KUKA KRL program: folge11.src, folge11.dat

--- folge11.src ---
&ACCESS RVP
&REL 1
&COMMENT bt2krl vw-ks24 production Folge 11 plan 16#A1BE
DEF FOLGE11()
   ; Generated by bt2krl 0.1.0 from bt2plc plan bt_1792156523_scene_fit (cell scene_fit), PLAN_ID 16#A1BE
   ; Robot robot1 (R1), controller robot1, model unknown, joint mapping identity
   ; Profile vw-ks24 (VW KS24 / TPVW 8.1.8).
   ; Do not edit: regenerate with bt2krl (plain KRL, no inline forms).
   ; Production Folge: 3 ops; per op: P_PktNr_SPS, interlock request + MAKRO20 handshake, motion (exact stop at the end), hold, interlock release
   ; The VW tech package does the Folge handshake (cell.src, AUE_INIT/WAIT/END).
   ;FOLD AUE INIT
      VW(#VW_AUE_INIT,TRUE)
      PENTER:
      INTERRUPT DECL 10 WHEN $CYCFLAG[254]==FALSE DO VW(#FB_STOP,TRUE)
      INTERRUPT ON 10
      INT10=TRUE
   ;ENDFOLD
   ;FOLD VWP0 P0 10 PCT
      ; P0 = home: VW_INIT runs BAS(#INITMOV); AUE_WAIT later sets $H_POS here
      VW(#VW_INIT,TRUE)
      VW_USR_R (#USR_INIT)
      BAS(#VEL_PTP,10)
      $APO.CPTP=100
      PTP P0
      $OUT[15]=TRUE ; PF0 Grundstellung
      ; MAKRO0 RUECKSETZEN_EA: resets A33-A96 (also the tool releases)
      SEL_RES=SELECT(#MAKRO,0,TRUE,,,,,FALSE)
   ;ENDFOLD
   ;FOLD VWAUEWAIT
      VW(#VW_AUE_WAIT,TRUE )
      IF N_VW==TRUE THEN
         GOTO PEXIT
      ENDIF
   ;ENDFOLD
   ;FOLD VWSTART 16#00000003
      ; release every interlock this robot uses: IL01=V1 IL02=V2
      $OUT[15]=FALSE ; PF0 off
      ; MAKRO50 Ini Merker: the cyclic flags of the driving conditions
      SEL_RES=SELECT(#MAKRO,50,TRUE,,,,,FALSE)
      $OUT[41]=TRUE ; release V1
      $OUT[42]=TRUE ; release V2
   ;ENDFOLD
   ;FOLD VWFB 16#00000000
      VALCYCFL30=$CYCFLAG[254]
      $CYCFLAG[254]=($CYCFLAG[30]) AND $CYCFLAG[255] OR ($TIMER[61]<0)
      VW(#FB_CHECK,TRUE)
   ;ENDFOLD
   ;FOLD OP 1 W02 MASK 16#00000001
      ; zones IL01
      P_PktNr_SPS=1
      ;FOLD VWLOCK 16#00000001
         ; enter IL01=V1
         $OUT[81]=TRUE ; request V1
         ; MAKRO20 semantics, inline for these interlocks only
         $OUT[41]=$OUT[41] OR $OUT[81]
         ; PLC grant of the request
         $LOOP_MSG[]="E81"
         $LOOP_CONT=TRUE
         WAIT FOR ($IN[81]) OR (NOT $LOOP_CONT AND ($MODE_OP<>#EX))
         $LOOP_MSG[]="                                                                                                                                "
         ; partner release
         $LOOP_MSG[]="E41"
         $LOOP_CONT=TRUE
         WAIT FOR ($IN[41]) OR (NOT $LOOP_CONT AND ($MODE_OP<>#EX))
         $LOOP_MSG[]="                                                                                                                                "
         $OUT[41]=FALSE ; occupied
         $OUT[81]=FALSE
      ;ENDFOLD
      ;FOLD VWFB 16#00000001
         VALCYCFL30=$CYCFLAG[254]
         $CYCFLAG[254]=($CYCFLAG[30] AND $IN[41]) AND $CYCFLAG[255] OR ($TIMER[61]<0)
         VW(#FB_CHECK,TRUE)
      ;ENDFOLD
      BAS(#VEL_PTP,3)
      PTP P1 C_PTP
      BAS(#VEL_PTP,5)
      PTP P2 C_PTP
      BAS(#VEL_PTP,8)
      PTP P3 C_PTP
      BAS(#VEL_PTP,11)
      PTP P4 C_PTP
      BAS(#VEL_PTP,13)
      PTP P5 C_PTP
      BAS(#VEL_PTP,12)
      PTP P6 C_PTP
      BAS(#VEL_PTP,9)
      PTP P7 C_PTP
      BAS(#VEL_PTP,7)
      PTP P8 C_PTP
      BAS(#VEL_PTP,5)
      PTP P9 C_PTP
      BAS(#VEL_PTP,2)
      PTP P10 C_PTP
      BAS(#VEL_PTP,6)
      PTP P11 C_PTP
      BAS(#VEL_PTP,8)
      PTP P12 C_PTP
      BAS(#VEL_PTP,3)
      PTP P13
      WAIT SEC 0.5 ; hold
      ;FOLD VWUNLOCK 16#00000001
         ; leave IL01=V1
         $OUT[41]=TRUE ; release V1
      ;ENDFOLD
      ;FOLD VWFB 16#00000000
         VALCYCFL30=$CYCFLAG[254]
         $CYCFLAG[254]=($CYCFLAG[30]) AND $CYCFLAG[255] OR ($TIMER[61]<0)
         VW(#FB_CHECK,TRUE)
      ;ENDFOLD
      WAIT SEC 0.1 ; step dwell
   ;ENDFOLD
   ;FOLD OP 2 W04 MASK 16#00000002
      ; zones IL02
      P_PktNr_SPS=2
      ;FOLD VWLOCK 16#00000002
         ; enter IL02=V2
         $OUT[82]=TRUE ; request V2
         ; MAKRO20 semantics, inline for these interlocks only
         $OUT[42]=$OUT[42] OR $OUT[82]
         ; PLC grant of the request
         $LOOP_MSG[]="E82"
         $LOOP_CONT=TRUE
         WAIT FOR ($IN[82]) OR (NOT $LOOP_CONT AND ($MODE_OP<>#EX))
         $LOOP_MSG[]="                                                                                                                                "
         ; partner release
         $LOOP_MSG[]="E42"
         $LOOP_CONT=TRUE
         WAIT FOR ($IN[42]) OR (NOT $LOOP_CONT AND ($MODE_OP<>#EX))
         $LOOP_MSG[]="                                                                                                                                "
         $OUT[42]=FALSE ; occupied
         $OUT[82]=FALSE
      ;ENDFOLD
      ;FOLD VWFB 16#00000002
         VALCYCFL30=$CYCFLAG[254]
         $CYCFLAG[254]=($CYCFLAG[30] AND $IN[42]) AND $CYCFLAG[255] OR ($TIMER[61]<0)
         VW(#FB_CHECK,TRUE)
      ;ENDFOLD
      BAS(#VEL_PTP,4)
      PTP P14 C_PTP
      PTP P15 C_PTP
      BAS(#VEL_PTP,10)
      PTP P16 C_PTP
      BAS(#VEL_PTP,13)
      PTP P17 C_PTP
      BAS(#VEL_PTP,11)
      PTP P18 C_PTP
      BAS(#VEL_PTP,7)
      PTP P19 C_PTP
      BAS(#VEL_PTP,3)
      PTP P20 C_PTP
      BAS(#VEL_PTP,6)
      PTP P21 C_PTP
      BAS(#VEL_PTP,8)
      PTP P22 C_PTP
      BAS(#VEL_PTP,3)
      PTP P23
      WAIT SEC 0.5 ; hold
      ;FOLD VWUNLOCK 16#00000002
         ; leave IL02=V2
         $OUT[42]=TRUE ; release V2
      ;ENDFOLD
      ;FOLD VWFB 16#00000000
         VALCYCFL30=$CYCFLAG[254]
         $CYCFLAG[254]=($CYCFLAG[30]) AND $CYCFLAG[255] OR ($TIMER[61]<0)
         VW(#FB_CHECK,TRUE)
      ;ENDFOLD
      WAIT SEC 0.1 ; step dwell
   ;ENDFOLD
   ;FOLD OP 3 HOME MASK 16#00000001
      ; zones IL01
      P_PktNr_SPS=3
      ;FOLD VWLOCK 16#00000001
         ; enter IL01=V1
         $OUT[81]=TRUE ; request V1
         ; MAKRO20 semantics, inline for these interlocks only
         $OUT[41]=$OUT[41] OR $OUT[81]
         ; PLC grant of the request
         $LOOP_MSG[]="E81"
         $LOOP_CONT=TRUE
         WAIT FOR ($IN[81]) OR (NOT $LOOP_CONT AND ($MODE_OP<>#EX))
         $LOOP_MSG[]="                                                                                                                                "
         ; partner release
         $LOOP_MSG[]="E41"
         $LOOP_CONT=TRUE
         WAIT FOR ($IN[41]) OR (NOT $LOOP_CONT AND ($MODE_OP<>#EX))
         $LOOP_MSG[]="                                                                                                                                "
         $OUT[41]=FALSE ; occupied
         $OUT[81]=FALSE
      ;ENDFOLD
      ;FOLD VWFB 16#00000001
         VALCYCFL30=$CYCFLAG[254]
         $CYCFLAG[254]=($CYCFLAG[30] AND $IN[41]) AND $CYCFLAG[255] OR ($TIMER[61]<0)
         VW(#FB_CHECK,TRUE)
      ;ENDFOLD
      BAS(#VEL_PTP,5)
      PTP P24 C_PTP
      BAS(#VEL_PTP,2)
      PTP P25 C_PTP
      BAS(#VEL_PTP,6)
      PTP P26 C_PTP
      BAS(#VEL_PTP,9)
      PTP P27 C_PTP
      BAS(#VEL_PTP,12)
      PTP P28 C_PTP
      BAS(#VEL_PTP,15)
      PTP P29 C_PTP
      BAS(#VEL_PTP,18)
      PTP P30 C_PTP
      BAS(#VEL_PTP,17)
      PTP P31 C_PTP
      BAS(#VEL_PTP,14)
      PTP P32 C_PTP
      BAS(#VEL_PTP,11)
      PTP P33 C_PTP
      BAS(#VEL_PTP,6)
      PTP P34 C_PTP
      BAS(#VEL_PTP,2)
      PTP P35
      ;FOLD VWMAKRO 15
         ; Gesamtfertigmeldung
         SEL_RES=SELECT(#MAKRO,15,TRUE,,,,,FALSE)
      ;ENDFOLD
      ;FOLD VWUNLOCK 16#00000001
         ; leave IL01=V1
         $OUT[41]=TRUE ; release V1
      ;ENDFOLD
      ;FOLD VWFB 16#00000000
         VALCYCFL30=$CYCFLAG[254]
         $CYCFLAG[254]=($CYCFLAG[30]) AND $CYCFLAG[255] OR ($TIMER[61]<0)
         VW(#FB_CHECK,TRUE)
      ;ENDFOLD
      WAIT SEC 0.1 ; step dwell
   ;ENDFOLD
   P_PktNr_SPS=0
   ;FOLD AUE END
      VW(#VW_AUE_END,TRUE)
      GOTO PENTER
      PEXIT:
   ;ENDFOLD
END

--- folge11.dat ---
&ACCESS RVP
&REL 1
&COMMENT bt2krl vw-ks24 data Folge 11 plan 16#A1BE
DEFDAT FOLGE11
   ; Generated by bt2krl 0.1.0 from bt2plc plan bt_1792156523_scene_fit (cell scene_fit), PLAN_ID 16#A1BE
   ; Robot robot1 (R1), controller robot1, model unknown, joint mapping identity
   ; Profile vw-ks24 (VW KS24 / TPVW 8.1.8).
   ; Do not edit: regenerate with bt2krl (plain KRL, no inline forms).
   EXT BAS (BAS_COMMAND :IN,REAL :IN )
   ; interface to the VW standard routines (as every VW Folge .dat declares them)
   EXT VW (VW_COMMAND :IN,BOOL :IN,REAL :IN,REAL :IN,REAL :IN,REAL :IN,BOOL :IN,E6POS :IN )
   EXT VW_USR_R (VW_USER_CMD :IN,INT :IN,REAL :IN,REAL :IN,REAL :IN,REAL :IN,REAL :IN,REAL :IN,BOOL :IN )
   EXTFCT INT SELECT (SUBTYPE :IN,INT :IN,BOOL :IN,ARI_TYP :IN,INT :IN,BOOL_TYP :IN,INT :IN,BOOL :IN)
   DECL AXIS P0={A1 45.0,A2 -90.0,A3 90.0,A4 0.0,A5 0.0,A6 0.0}
   DECL AXIS P1={A1 43.6012,A2 -89.7676,A3 90.0033,A4 0.0,A5 1.8605,A6 -0.3507}
   DECL AXIS P2={A1 41.9543,A2 -89.4939,A3 90.0071,A4 0.0,A5 4.051,A6 -0.7636}
   DECL AXIS P3={A1 37.1038,A2 -88.6879,A3 90.0185,A4 0.0,A5 10.5026,A6 -1.9796}
   DECL AXIS P4={A1 26.9514,A2 -87.001,A3 90.0423,A4 0.0,A5 24.006,A6 -4.5249}
   DECL AXIS P5={A1 6.8724,A2 -83.6646,A3 90.0893,A4 0.0,A5 50.7127,A6 -9.5588}
   DECL AXIS P6={A1 -4.0921,A2 -81.8426,A3 90.115,A4 0.0,A5 65.2964,A6 -12.3077}
   DECL AXIS P7={A1 -9.8225,A2 -80.8905,A3 90.1284,A4 0.0,A5 72.9183,A6 -13.7444}
   DECL AXIS P8={A1 -12.0109,A2 -80.5268,A3 90.1336,A4 0.0,A5 75.829,A6 -14.293}
   DECL AXIS P9={A1 -14.6956,A2 -80.0807,A3 90.1398,A4 0.0,A5 79.3999,A6 -14.9661}
   DECL AXIS P10={A1 -15.0566,A2 -80.0207,A3 90.1407,A4 0.0,A5 79.88,A6 -15.0566}
   DECL AXIS P11={A1 -15.0566,A2 -79.875,A3 90.7142,A4 0.0,A5 79.1607,A6 -15.0566}
   DECL AXIS P12={A1 -15.0566,A2 -79.6592,A3 91.5498,A4 0.0,A5 78.1094,A6 -15.0566}
   DECL AXIS P13={A1 -15.0566,A2 -78.7933,A3 94.228,A4 0.0,A5 74.5653,A6 -15.0566}
   DECL AXIS P14={A1 -15.0374,A2 -79.913,A3 90.5893,A4 0.0,A5 79.3237,A6 -15.0374}
   DECL AXIS P15={A1 -13.7654,A2 -80.0274,A3 90.142,A4 0.0,A5 79.8854,A6 -13.7654}
   DECL AXIS P16={A1 -9.2939,A2 -80.052,A3 90.1253,A4 0.0,A5 79.9267,A6 -9.2939}
   DECL AXIS P17={A1 8.1168,A2 -80.1118,A3 90.221,A4 0.0,A5 79.8908,A6 8.1168}
   DECL AXIS P18={A1 11.5499,A2 -80.1218,A3 90.2471,A4 0.0,A5 79.8747,A6 11.5498}
   DECL AXIS P19={A1 13.8795,A2 -80.1284,A3 90.2658,A4 0.0,A5 79.8625,A6 13.8794}
   DECL AXIS P20={A1 14.7377,A2 -80.1307,A3 90.273,A4 0.0,A5 79.8577,A6 14.7377}
   DECL AXIS P21={A1 14.7377,A2 -79.9847,A3 90.8466,A4 0.0,A5 79.1381,A6 14.7377}
   DECL AXIS P22={A1 14.7377,A2 -79.7685,A3 91.6823,A4 0.0,A5 78.0862,A6 14.7377}
   DECL AXIS P23={A1 14.7377,A2 -78.9012,A3 94.361,A4 0.0,A5 74.5402,A6 14.7377}
   DECL AXIS P24={A1 14.7377,A2 -79.9556,A3 90.9835,A4 0.0,A5 78.9721,A6 14.7377}
   DECL AXIS P25={A1 15.0076,A2 -80.0451,A3 90.9747,A4 0.0,A5 78.2679,A6 14.6063}
   DECL AXIS P26={A1 15.7755,A2 -80.3,A3 90.9498,A4 0.0,A5 76.2638,A6 14.2323}
   DECL AXIS P27={A1 16.9794,A2 -80.6996,A3 90.9106,A4 0.0,A5 73.1223,A6 13.646}
   DECL AXIS P28={A1 18.5568,A2 -81.2232,A3 90.8594,A4 0.0,A5 69.0058,A6 12.8778}
   DECL AXIS P29={A1 22.5835,A2 -82.5597,A3 90.7285,A4 0.0,A5 58.4978,A6 10.9168}
   DECL AXIS P30={A1 34.8296,A2 -86.6243,A3 90.3305,A4 0.0,A5 26.5407,A6 4.953}
   DECL AXIS P31={A1 39.2921,A2 -88.1055,A3 90.1855,A4 0.0,A5 14.8953,A6 2.7797}
   DECL AXIS P32={A1 41.1809,A2 -88.7324,A3 90.1241,A4 0.0,A5 9.9663,A6 1.8599}
   DECL AXIS P33={A1 43.9622,A2 -89.6555,A3 90.0337,A4 0.0,A5 2.7082,A6 0.5054}
   DECL AXIS P34={A1 44.7302,A2 -89.9104,A3 90.0088,A4 0.0,A5 0.7041,A6 0.1314}
   DECL AXIS P35={A1 45.0,A2 -90.0,A3 90.0,A4 0.0,A5 0.0,A6 0.0}
ENDDAT
